Staubli VAL3: pickAndPlace.pgx

program pickAndPlace()
// Lab2A Level 3 - shared manual simulation / physical cycle
begin

  // Pick from the selected ramp.
  vacuumOn = false
  blowOn = false

  movej(pickApproach[materialType], vacuumTool, moveSpeed)
  waitEndMove()

  movel(jointToPoint(vacuumTool, world, pickPose[materialType]), vacuumTool, moveSpeed)
  waitEndMove()

  vacuumOn = true
  cycleStep = 60
  putln("60 - Picking part: waiting for vacuum confirmation (partOnTool=true)")
  wait(partOnTool == true)

  movel(jointToPoint(vacuumTool, world, pickApproach[materialType]), vacuumTool, moveSpeed)
  waitEndMove()

  // Transfer and release at the selected destination.
  movej(placeApproach[placeIndex], vacuumTool, moveSpeed)
  waitEndMove()

  movel(jointToPoint(vacuumTool, world, placePose[placeIndex]), vacuumTool, moveSpeed)
  waitEndMove()

  vacuumOn = false
  blowOn = true
  delay(0.3)
  blowOn = false
  cycleStep = 70
  putln("70 - Releasing part: waiting for release confirmation (partOnTool=false)")
  wait(partOnTool == false)

  // Withdraw and return home.
  movel(jointToPoint(vacuumTool, world, placeApproach[placeIndex]), vacuumTool, moveSpeed)
  waitEndMove()

  movej(homePose, vacuumTool, moveSpeed)
  waitEndMove()

end
